// TIA Portal V20 export
// export: Created 2026-03-20T09:31:01.8595243Z, ExportSetting WithDefaults, DisplayName Totally Integrated Automation Portal, DisplayVersion V20, DisplayName TIA Portal Openness, DisplayVersion V20, DisplayName TIA Portal Version Control Interface, DisplayVersion V20, DisplayName TIA Portal Test Suite Advanced, DisplayVersion V20, DisplayName STEP 7 Professional, DisplayVersion V20, DisplayName STEP 7 Safety, DisplayVersion V20, DisplayName WinCC Basic/Comfort/Advanced, DisplayVersion V20
FUNCTION_BLOCK "LifterSeq_79bef3"   // FB1, LAD
VERSION : 0.1
// stored: AutoNumber true, IsIECCheckEnabled false, UDAEnableTagReadback false
   VAR_INPUT
      iArea_Clear : Bool;
      iAutoRunning : Bool;
      iLifter_Down_over : Bool;
      iLifter_Up_over : Bool;
      iNext_Stan_RTR : Bool;
      iOTS_from_Prevous_STN : Bool;
      iReset_fault : Bool;
      iSstMode : Bool;
      iSstPB : Bool;
   END_VAR
   VAR_OUTPUT
      qLifter_DOWN_CMD : Bool;
      qLifter_UP_CMD : Bool;
   END_VAR
   VAR DB_SPECIFIC
      StateNo : Int;
      s10_WaitForStart : Bool;
      s10_WaitForStart_T1 : Bool;
      s11_ChkPalletPrsnt : Bool;
      s11_ChkPalletPrsnt_T1 : Bool;
      s11_ChkPalletPrsnt_T2 : Bool;
      s12_WaitAreaClear : Bool;
      s12_WaitAreaClear_T1 : Bool;
      s14_WaitLifterDown : Bool;
      s14_WaitLifterDown_T1 : Bool;
      s15_WaitNextStnRdy : Bool;
      s15_WaitNextStnRdy_T1 : Bool;
      s16_WaitPalletAbsnt : Bool;
      s16_WaitPalletAbsnt_T1 : Bool;
      s17_WaitAreaClear : Bool;
      s17_WaitAreaClear_T1 : Bool;
      s18_WaitLifterUp : Bool;
      s18_WaitLifterUp_T1 : Bool;
      sSst : Bool;
      sSstPulse : Bool;
      sSstRise : Bool;
      sStWtResetRel : Bool;
      sStWtResetRel_T1 : Bool;
   END_VAR
   VAR_TEMP
      tOne : Bool;
   END_VAR
   VAR_TEMP   // added for the SCL form of the ladder/FBD networks
      _w1 : Bool;
   END_VAR
BEGIN

REGION Network 1
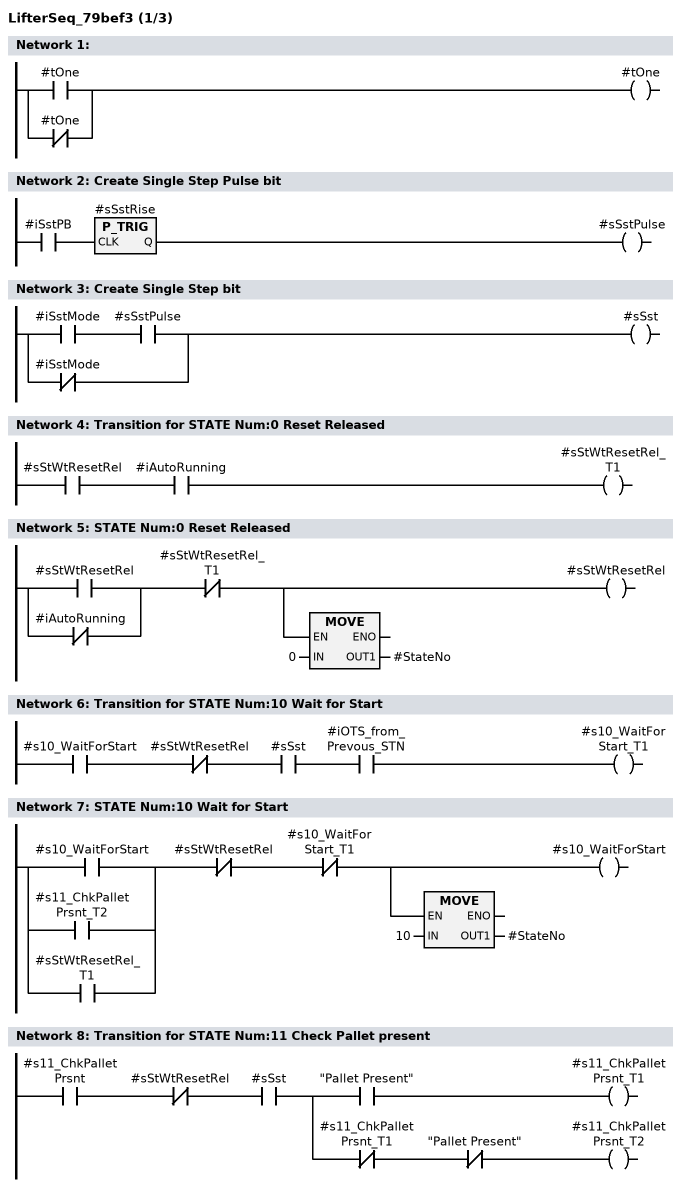
   RUNG wire#powerrail
      Contact( #tOne )
      wire#w1
      Coil( #tOne )
   END_RUNG
   RUNG wire#powerrail
      I_Contact( #tOne )
   END_RUNG wire#w1
   // the same network as SCL:
   #tOne := #tOne OR NOT #tOne;
END_REGION

REGION Network 2: Create Single Step Pulse bit
   RUNG wire#powerrail
      Contact( #iSstPB )
      P_Trig( #sSstRise )
      Coil( #sSstPulse )
   END_RUNG
   // the same network as SCL:
   #_w1 := #iSstPB AND NOT #sSstRise;   // rising edge
   #sSstRise := #iSstPB;
   #sSstPulse := #_w1;
END_REGION

REGION Network 3: Create Single Step bit
   RUNG wire#powerrail
      Contact( #iSstMode )
      Contact( #sSstPulse )
      wire#w1
      Coil( #sSst )
   END_RUNG
   RUNG wire#powerrail
      I_Contact( #iSstMode )
   END_RUNG wire#w1
   // the same network as SCL:
   #sSst := (#iSstMode AND #sSstPulse) OR NOT #iSstMode;
END_REGION

REGION Network 4: Transition for STATE Num:0 Reset Released
   RUNG wire#powerrail
      Contact( #sStWtResetRel )
      Contact( #iAutoRunning )
      Coil( #sStWtResetRel_T1 )
   END_RUNG
   // the same network as SCL:
   #sStWtResetRel_T1 := #sStWtResetRel AND #iAutoRunning;
END_REGION

REGION Network 5: STATE Num:0 Reset Released
   RUNG wire#powerrail
      Contact( #sStWtResetRel )
      wire#w1
      I_Contact( #sStWtResetRel_T1 )
      wire#w2
      Coil( #sStWtResetRel )
   END_RUNG
   RUNG wire#powerrail
      I_Contact( #iAutoRunning )
   END_RUNG wire#w1
   RUNG wire#w2
      { S7_GenerateENO := "TRUE" } Move(in := 0, out1 => #StateNo)
   END_RUNG
   // the same network as SCL:
   #sStWtResetRel := (#sStWtResetRel OR NOT #iAutoRunning) AND NOT #sStWtResetRel_T1;
   IF #sStWtResetRel THEN #StateNo := 0; END_IF;
END_REGION

REGION Network 6: Transition for STATE Num:10 Wait for Start
   RUNG wire#powerrail
      Contact( #s10_WaitForStart )
      I_Contact( #sStWtResetRel )
      Contact( #sSst )
      Contact( #iOTS_from_Prevous_STN )
      Coil( #s10_WaitForStart_T1 )
   END_RUNG
   // the same network as SCL:
   #s10_WaitForStart_T1 := #s10_WaitForStart AND NOT #sStWtResetRel AND #sSst AND #iOTS_from_Prevous_STN;
END_REGION

REGION Network 7: STATE Num:10 Wait for Start
   RUNG wire#powerrail
      Contact( #s10_WaitForStart )
      wire#w1
      I_Contact( #sStWtResetRel )
      I_Contact( #s10_WaitForStart_T1 )
      wire#w2
      Coil( #s10_WaitForStart )
   END_RUNG
   RUNG wire#powerrail
      Contact( #s11_ChkPalletPrsnt_T2 )
   END_RUNG wire#w1
   RUNG wire#powerrail
      Contact( #sStWtResetRel_T1 )
   END_RUNG wire#w1
   RUNG wire#w2
      { S7_GenerateENO := "TRUE" } Move(in := 10, out1 => #StateNo)
   END_RUNG
   // the same network as SCL:
   #s10_WaitForStart := (#s10_WaitForStart OR #s11_ChkPalletPrsnt_T2 OR #sStWtResetRel_T1) AND NOT #sStWtResetRel AND NOT #s10_WaitForStart_T1;
   IF #s10_WaitForStart THEN #StateNo := 10; END_IF;
END_REGION

REGION Network 8: Transition for STATE Num:11 Check Pallet present
   RUNG wire#powerrail
      Contact( #s11_ChkPalletPrsnt )
      I_Contact( #sStWtResetRel )
      Contact( #sSst )
      wire#w1
      Contact( "Pallet Present" )
      Coil( #s11_ChkPalletPrsnt_T1 )
   END_RUNG
   RUNG wire#w1
      I_Contact( #s11_ChkPalletPrsnt_T1 )
      I_Contact( "Pallet Present" )
      Coil( #s11_ChkPalletPrsnt_T2 )
   END_RUNG
   // the same network as SCL:
   #_w1 := #s11_ChkPalletPrsnt AND NOT #sStWtResetRel AND #sSst;
   #s11_ChkPalletPrsnt_T1 := #_w1 AND "Pallet Present";
   #s11_ChkPalletPrsnt_T2 := #_w1 AND NOT #s11_ChkPalletPrsnt_T1 AND NOT "Pallet Present";
END_REGION

REGION Network 9: STATE Num:11 Check Pallet present
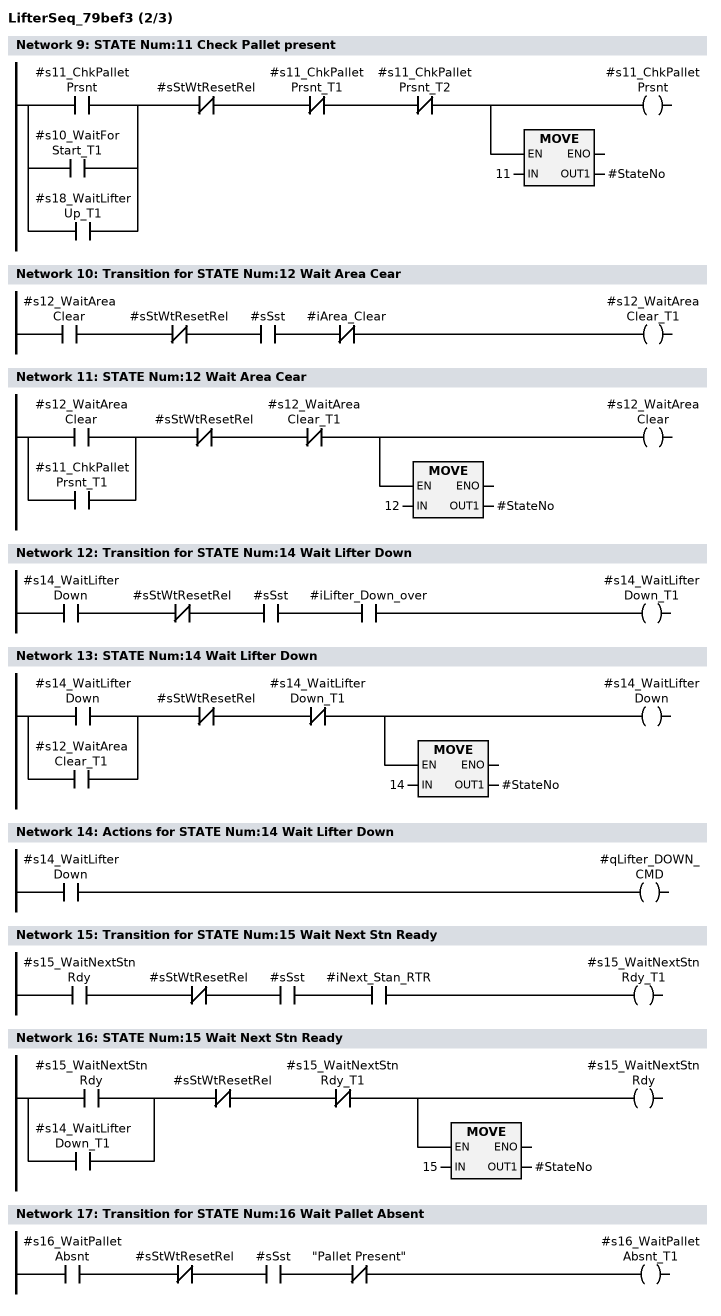
   RUNG wire#powerrail
      Contact( #s11_ChkPalletPrsnt )
      wire#w1
      I_Contact( #sStWtResetRel )
      I_Contact( #s11_ChkPalletPrsnt_T1 )
      I_Contact( #s11_ChkPalletPrsnt_T2 )
      wire#w2
      Coil( #s11_ChkPalletPrsnt )
   END_RUNG
   RUNG wire#powerrail
      Contact( #s10_WaitForStart_T1 )
   END_RUNG wire#w1
   RUNG wire#powerrail
      Contact( #s18_WaitLifterUp_T1 )
   END_RUNG wire#w1
   RUNG wire#w2
      { S7_GenerateENO := "TRUE" } Move(in := 11, out1 => #StateNo)
   END_RUNG
   // the same network as SCL:
   #s11_ChkPalletPrsnt := (#s11_ChkPalletPrsnt OR #s10_WaitForStart_T1 OR #s18_WaitLifterUp_T1) AND NOT #sStWtResetRel AND NOT #s11_ChkPalletPrsnt_T1 AND NOT #s11_ChkPalletPrsnt_T2;
   IF #s11_ChkPalletPrsnt THEN #StateNo := 11; END_IF;
END_REGION

REGION Network 10: Transition for STATE Num:12 Wait Area Cear
   RUNG wire#powerrail
      Contact( #s12_WaitAreaClear )
      I_Contact( #sStWtResetRel )
      Contact( #sSst )
      I_Contact( #iArea_Clear )
      Coil( #s12_WaitAreaClear_T1 )
   END_RUNG
   // the same network as SCL:
   #s12_WaitAreaClear_T1 := #s12_WaitAreaClear AND NOT #sStWtResetRel AND #sSst AND NOT #iArea_Clear;
END_REGION

REGION Network 11: STATE Num:12 Wait Area Cear
   RUNG wire#powerrail
      Contact( #s12_WaitAreaClear )
      wire#w1
      I_Contact( #sStWtResetRel )
      I_Contact( #s12_WaitAreaClear_T1 )
      wire#w2
      Coil( #s12_WaitAreaClear )
   END_RUNG
   RUNG wire#powerrail
      Contact( #s11_ChkPalletPrsnt_T1 )
   END_RUNG wire#w1
   RUNG wire#w2
      { S7_GenerateENO := "TRUE" } Move(in := 12, out1 => #StateNo)
   END_RUNG
   // the same network as SCL:
   #s12_WaitAreaClear := (#s12_WaitAreaClear OR #s11_ChkPalletPrsnt_T1) AND NOT #sStWtResetRel AND NOT #s12_WaitAreaClear_T1;
   IF #s12_WaitAreaClear THEN #StateNo := 12; END_IF;
END_REGION

REGION Network 12: Transition for STATE Num:14 Wait Lifter Down
   RUNG wire#powerrail
      Contact( #s14_WaitLifterDown )
      I_Contact( #sStWtResetRel )
      Contact( #sSst )
      Contact( #iLifter_Down_over )
      Coil( #s14_WaitLifterDown_T1 )
   END_RUNG
   // the same network as SCL:
   #s14_WaitLifterDown_T1 := #s14_WaitLifterDown AND NOT #sStWtResetRel AND #sSst AND #iLifter_Down_over;
END_REGION

REGION Network 13: STATE Num:14 Wait Lifter Down
   RUNG wire#powerrail
      Contact( #s14_WaitLifterDown )
      wire#w1
      I_Contact( #sStWtResetRel )
      I_Contact( #s14_WaitLifterDown_T1 )
      wire#w2
      Coil( #s14_WaitLifterDown )
   END_RUNG
   RUNG wire#powerrail
      Contact( #s12_WaitAreaClear_T1 )
   END_RUNG wire#w1
   RUNG wire#w2
      { S7_GenerateENO := "TRUE" } Move(in := 14, out1 => #StateNo)
   END_RUNG
   // the same network as SCL:
   #s14_WaitLifterDown := (#s14_WaitLifterDown OR #s12_WaitAreaClear_T1) AND NOT #sStWtResetRel AND NOT #s14_WaitLifterDown_T1;
   IF #s14_WaitLifterDown THEN #StateNo := 14; END_IF;
END_REGION

REGION Network 14: Actions for STATE Num:14 Wait Lifter Down
   RUNG wire#powerrail
      Contact( #s14_WaitLifterDown )
      Coil( #qLifter_DOWN_CMD )
   END_RUNG
   // the same network as SCL:
   #qLifter_DOWN_CMD := #s14_WaitLifterDown;
END_REGION

REGION Network 15: Transition for STATE Num:15 Wait Next Stn Ready
   RUNG wire#powerrail
      Contact( #s15_WaitNextStnRdy )
      I_Contact( #sStWtResetRel )
      Contact( #sSst )
      Contact( #iNext_Stan_RTR )
      Coil( #s15_WaitNextStnRdy_T1 )
   END_RUNG
   // the same network as SCL:
   #s15_WaitNextStnRdy_T1 := #s15_WaitNextStnRdy AND NOT #sStWtResetRel AND #sSst AND #iNext_Stan_RTR;
END_REGION

REGION Network 16: STATE Num:15 Wait Next Stn Ready
   RUNG wire#powerrail
      Contact( #s15_WaitNextStnRdy )
      wire#w1
      I_Contact( #sStWtResetRel )
      I_Contact( #s15_WaitNextStnRdy_T1 )
      wire#w2
      Coil( #s15_WaitNextStnRdy )
   END_RUNG
   RUNG wire#powerrail
      Contact( #s14_WaitLifterDown_T1 )
   END_RUNG wire#w1
   RUNG wire#w2
      { S7_GenerateENO := "TRUE" } Move(in := 15, out1 => #StateNo)
   END_RUNG
   // the same network as SCL:
   #s15_WaitNextStnRdy := (#s15_WaitNextStnRdy OR #s14_WaitLifterDown_T1) AND NOT #sStWtResetRel AND NOT #s15_WaitNextStnRdy_T1;
   IF #s15_WaitNextStnRdy THEN #StateNo := 15; END_IF;
END_REGION

REGION Network 17: Transition for STATE Num:16 Wait Pallet Absent
   RUNG wire#powerrail
      Contact( #s16_WaitPalletAbsnt )
      I_Contact( #sStWtResetRel )
      Contact( #sSst )
      I_Contact( "Pallet Present" )
      Coil( #s16_WaitPalletAbsnt_T1 )
   END_RUNG
   // the same network as SCL:
   #s16_WaitPalletAbsnt_T1 := #s16_WaitPalletAbsnt AND NOT #sStWtResetRel AND #sSst AND NOT "Pallet Present";
END_REGION

REGION Network 18: STATE Num:16 Wait Pallet Absent
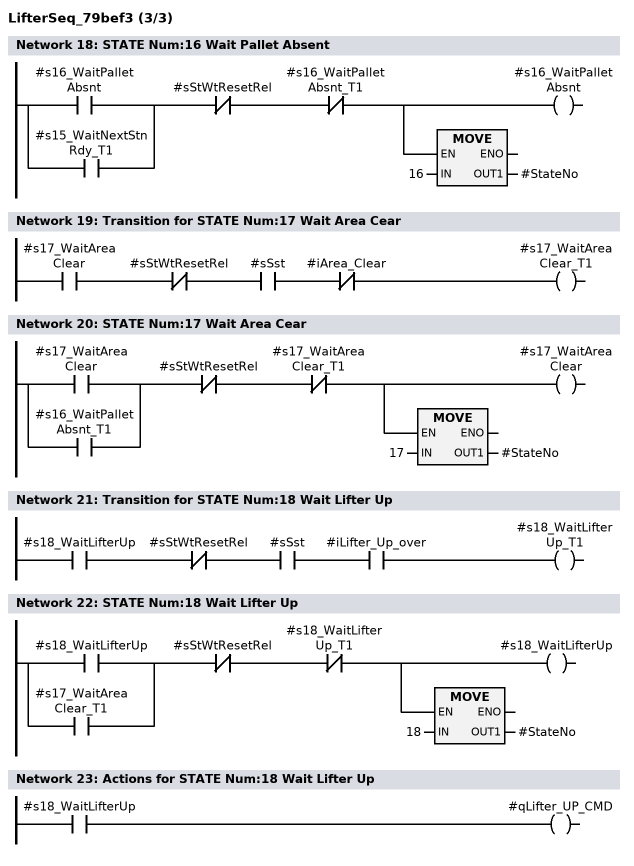
   RUNG wire#powerrail
      Contact( #s16_WaitPalletAbsnt )
      wire#w1
      I_Contact( #sStWtResetRel )
      I_Contact( #s16_WaitPalletAbsnt_T1 )
      wire#w2
      Coil( #s16_WaitPalletAbsnt )
   END_RUNG
   RUNG wire#powerrail
      Contact( #s15_WaitNextStnRdy_T1 )
   END_RUNG wire#w1
   RUNG wire#w2
      { S7_GenerateENO := "TRUE" } Move(in := 16, out1 => #StateNo)
   END_RUNG
   // the same network as SCL:
   #s16_WaitPalletAbsnt := (#s16_WaitPalletAbsnt OR #s15_WaitNextStnRdy_T1) AND NOT #sStWtResetRel AND NOT #s16_WaitPalletAbsnt_T1;
   IF #s16_WaitPalletAbsnt THEN #StateNo := 16; END_IF;
END_REGION

REGION Network 19: Transition for STATE Num:17 Wait Area Cear
   RUNG wire#powerrail
      Contact( #s17_WaitAreaClear )
      I_Contact( #sStWtResetRel )
      Contact( #sSst )
      I_Contact( #iArea_Clear )
      Coil( #s17_WaitAreaClear_T1 )
   END_RUNG
   // the same network as SCL:
   #s17_WaitAreaClear_T1 := #s17_WaitAreaClear AND NOT #sStWtResetRel AND #sSst AND NOT #iArea_Clear;
END_REGION

REGION Network 20: STATE Num:17 Wait Area Cear
   RUNG wire#powerrail
      Contact( #s17_WaitAreaClear )
      wire#w1
      I_Contact( #sStWtResetRel )
      I_Contact( #s17_WaitAreaClear_T1 )
      wire#w2
      Coil( #s17_WaitAreaClear )
   END_RUNG
   RUNG wire#powerrail
      Contact( #s16_WaitPalletAbsnt_T1 )
   END_RUNG wire#w1
   RUNG wire#w2
      { S7_GenerateENO := "TRUE" } Move(in := 17, out1 => #StateNo)
   END_RUNG
   // the same network as SCL:
   #s17_WaitAreaClear := (#s17_WaitAreaClear OR #s16_WaitPalletAbsnt_T1) AND NOT #sStWtResetRel AND NOT #s17_WaitAreaClear_T1;
   IF #s17_WaitAreaClear THEN #StateNo := 17; END_IF;
END_REGION

REGION Network 21: Transition for STATE Num:18 Wait Lifter Up
   RUNG wire#powerrail
      Contact( #s18_WaitLifterUp )
      I_Contact( #sStWtResetRel )
      Contact( #sSst )
      Contact( #iLifter_Up_over )
      Coil( #s18_WaitLifterUp_T1 )
   END_RUNG
   // the same network as SCL:
   #s18_WaitLifterUp_T1 := #s18_WaitLifterUp AND NOT #sStWtResetRel AND #sSst AND #iLifter_Up_over;
END_REGION

REGION Network 22: STATE Num:18 Wait Lifter Up
   RUNG wire#powerrail
      Contact( #s18_WaitLifterUp )
      wire#w1
      I_Contact( #sStWtResetRel )
      I_Contact( #s18_WaitLifterUp_T1 )
      wire#w2
      Coil( #s18_WaitLifterUp )
   END_RUNG
   RUNG wire#powerrail
      Contact( #s17_WaitAreaClear_T1 )
   END_RUNG wire#w1
   RUNG wire#w2
      { S7_GenerateENO := "TRUE" } Move(in := 18, out1 => #StateNo)
   END_RUNG
   // the same network as SCL:
   #s18_WaitLifterUp := (#s18_WaitLifterUp OR #s17_WaitAreaClear_T1) AND NOT #sStWtResetRel AND NOT #s18_WaitLifterUp_T1;
   IF #s18_WaitLifterUp THEN #StateNo := 18; END_IF;
END_REGION

REGION Network 23: Actions for STATE Num:18 Wait Lifter Up
   RUNG wire#powerrail
      Contact( #s18_WaitLifterUp )
      Coil( #qLifter_UP_CMD )
   END_RUNG
   // the same network as SCL:
   #qLifter_UP_CMD := #s18_WaitLifterUp;
END_REGION
END_FUNCTION_BLOCK
